(* IEC 61131-3 sources: codesys-to-astra/tools/tests/fixtures/sample/tests/POUs/FB_F_Clamp_Test, 4 files *)

(* ---- FB_F_Clamp_Test.decl.st ---- *)
(*
    Назначение: тесты CfUnit для F_Clamp — граничные условия и перепутанные границы
    Автор: kr0nsch
    Версия: 1.0.0
    Документ: docs/TEST_REPORT.md
*)
FUNCTION_BLOCK FB_F_Clamp_Test EXTENDS CfUnit.FB_TestSuite
VAR
END_VAR

(* ---- SwappedLimits.method.decl.st ---- *)
METHOD PRIVATE SwappedLimits
VAR
    rResult : REAL;
END_VAR

(* ---- ValueBelowMin.method.decl.st ---- *)
METHOD PRIVATE ValueBelowMin
VAR
    rResult : REAL;
END_VAR

(* ---- ValueInsideRange.method.decl.st ---- *)
METHOD PRIVATE ValueInsideRange
VAR
    rResult : REAL;
END_VAR
